FUNCTION_BLOCK FB_CartonCell EXTENDS SPT_BaseTypes.FB_PackML_BaseModule
VAR
    Line : FB_ContinuousLine;
    LineEvents : FB_LineEvents;
    Devices : FB_CellDevices;
    Stations : ARRAY[1..5] OF FB_StrokeStation;
    ActiveStation : DINT;
    Finished : BOOL;
    Cartons : DINT;
    AirFault : BOOL;
    LowStock : BOOL;
    PreviousState : Tc3_PackML_V2.E_PMLState;
    ActingScans : INT;
    RequestSample : DINT;
    Acknowledged : DINT;
    Accepted : BOOL;
    StatusBuffer : ARRAY[0..105] OF DINT;
END_VAR

METHOD PROTECTED Initialize : BOOL
// User mode 4 keeps Idle and Complete for one-station commissioning.
CustomModes(eMode := 4, sName := 'Manual stroke', bDisableHeld := TRUE,
    bDisableSuspended := TRUE, bEnableUnitModeChangeStopped := TRUE);
Initialize := SUPER^.Initialize();
END_METHOD

METHOD RunScan
IF _InitComplete THEN
    CyclicLogic();
ELSE
    _InitComplete := Initialize();
END_IF
END_METHOD

METHOD CyclicLogic
// SPT can call this hook while Initialize is still on the stack.
IF NOT _InitComplete THEN RETURN; END_IF

IF _CurrentState <> PreviousState THEN
    ActingScans := 0;
    PreviousState := _CurrentState;
ELSE
    ActingScans := MIN(45, ActingScans + 1);
END_IF

// Sample once so a concurrent ADS write belongs entirely to one scan.
RequestSample := GVL_HMI.Request;
IF RequestSample <> Acknowledged THEN
    Accepted := ApplyCommand(RequestSample MOD 256);
    Acknowledged := RequestSample;
END_IF

Line.Clock((_CurrentState = Tc3_PackML_V2.E_PMLState.ePMLState_Execute) AND Line.Enabled AND (_CurrentMode = E_PMLUnitMode.ePMLUnitMode_Production));
SUPER^.CyclicLogic();
LineEvents(Occurrence := Line.Occurrence, Alarm := Line.Alarm, Jammed := Line.Jammed,
    Idle := _CurrentState = Tc3_PackML_V2.E_PMLState.ePMLState_Idle);
PublishStatus();
END_METHOD

METHOD PROTECTED Execute
IF Line.Enabled AND (_CurrentMode = E_PMLUnitMode.ePMLUnitMode_Production) THEN
    IF Line.Alarm = 0 THEN Line.Step(Devices.MissingSeal); END_IF
    IF Line.Alarm <> 0 THEN ChangeState(Tc3_PackML_V2.E_PMLCommand.ePMLCommand_Abort); END_IF
    RETURN;
END_IF
IF (ActiveStation < 1) OR (ActiveStation > 5) THEN RETURN; END_IF
IF Finished THEN
    StateComplete();
    RETURN;
END_IF

Stations[ActiveStation].Step();
IF _CurrentMode = E_PMLUnitMode.ePMLUnitMode_Production THEN
    Devices.ProcessStation(ActiveStation, Stations[ActiveStation].Phase);
END_IF

IF Stations[ActiveStation].Done AND
   ((_CurrentMode = E_PMLUnitMode.ePMLUnitMode_UserMode1) OR Devices.ReadyToLeave(ActiveStation)) THEN
    IF (_CurrentMode = E_PMLUnitMode.ePMLUnitMode_UserMode1) OR (ActiveStation = 5) THEN
        Finished := TRUE;
        IF _CurrentMode = E_PMLUnitMode.ePMLUnitMode_Production THEN
            IF Devices.FinishCarton() THEN
                Cartons := Cartons + 1;
            END_IF
        END_IF
        StateComplete();
    ELSIF Devices.IndexToNext(ActiveStation) THEN
        ActiveStation := ActiveStation + 1;
    END_IF
END_IF
END_METHOD

METHOD PROTECTED Resetting
VAR
    StationIndex : INT;
END_VAR
FOR StationIndex := 1 TO 5 DO
    Stations[StationIndex].ResetStation();
END_FOR
Devices.ResetDevices();
Line.ResetLine();
ActiveStation := 0;
Finished := FALSE;
IF (_CurrentState = PreviousState) AND (ActingScans >= 45) THEN
    StateComplete();
END_IF
END_METHOD

METHOD PROTECTED Clearing
IF (_CurrentState = PreviousState) AND (ActingScans >= 45) THEN
    StateComplete();
END_IF
END_METHOD

METHOD PROTECTED Starting
IF (_CurrentState = PreviousState) AND (ActingScans >= 45) THEN
    StateComplete();
END_IF
END_METHOD

METHOD PROTECTED Stopping
IF (_CurrentState = PreviousState) AND (ActingScans >= 45) THEN
    StateComplete();
END_IF
END_METHOD

METHOD PROTECTED Aborting
IF (_CurrentState = PreviousState) AND (ActingScans >= 45) THEN
    StateComplete();
END_IF
END_METHOD

METHOD PROTECTED Holding
IF (_CurrentState = PreviousState) AND (ActingScans >= 45) THEN
    StateComplete();
END_IF
END_METHOD

METHOD PROTECTED Unholding
IF (_CurrentState = PreviousState) AND (ActingScans >= 45) THEN
    StateComplete();
END_IF
END_METHOD

METHOD PROTECTED Suspending
IF (_CurrentState = PreviousState) AND (ActingScans >= 45) THEN
    StateComplete();
END_IF
END_METHOD

METHOD PROTECTED Unsuspending
IF (_CurrentState = PreviousState) AND (ActingScans >= 45) THEN
    StateComplete();
END_IF
END_METHOD

METHOD PROTECTED Completing
IF (_CurrentState = PreviousState) AND (ActingScans >= 45) THEN
    StateComplete();
END_IF
END_METHOD

METHOD PRIVATE ApplyCommand : BOOL
VAR_INPUT
    Code : DINT;
END_VAR
VAR
    IsManual : BOOL;
END_VAR
IsManual := _CurrentMode = E_PMLUnitMode.ePMLUnitMode_UserMode1;
CASE Code OF
    E_ConsoleCommand.Reset:
        IF NOT AirFault AND ((_CurrentState = Tc3_PackML_V2.E_PMLState.ePMLState_Stopped) OR (_CurrentState = Tc3_PackML_V2.E_PMLState.ePMLState_Complete)) THEN
            ChangeState(Tc3_PackML_V2.E_PMLCommand.ePMLCommand_Reset);
            ApplyCommand := TRUE;
        END_IF
    E_ConsoleCommand.Start:
        IF NOT IsManual AND (_CurrentState = Tc3_PackML_V2.E_PMLState.ePMLState_Idle) THEN
            Line.Timing := Line.Enabled;
            ActiveStation := SEL(Line.Enabled, 1, 0);
            ChangeState(Tc3_PackML_V2.E_PMLCommand.ePMLCommand_Start);
            ApplyCommand := TRUE;
        END_IF
    E_ConsoleCommand.Hold:
        IF NOT IsManual AND (_CurrentState = Tc3_PackML_V2.E_PMLState.ePMLState_Execute) THEN
            ChangeState(Tc3_PackML_V2.E_PMLCommand.ePMLCommand_Hold);
            ApplyCommand := TRUE;
        END_IF
    E_ConsoleCommand.Unhold:
        IF _CurrentState = Tc3_PackML_V2.E_PMLState.ePMLState_Held THEN
            ChangeState(Tc3_PackML_V2.E_PMLCommand.ePMLCommand_Unhold);
            ApplyCommand := TRUE;
        END_IF
    E_ConsoleCommand.Suspend:
        IF NOT IsManual AND (_CurrentState = Tc3_PackML_V2.E_PMLState.ePMLState_Execute) THEN
            ChangeState(Tc3_PackML_V2.E_PMLCommand.ePMLCommand_Suspend);
            ApplyCommand := TRUE;
        END_IF
    E_ConsoleCommand.Unsuspend:
        IF _CurrentState = Tc3_PackML_V2.E_PMLState.ePMLState_Suspended THEN
            ChangeState(Tc3_PackML_V2.E_PMLCommand.ePMLCommand_Unsuspend);
            ApplyCommand := TRUE;
        END_IF
    E_ConsoleCommand.Stop:
        IF (_CurrentState <> Tc3_PackML_V2.E_PMLState.ePMLState_Undefined) AND
            (_CurrentState <> Tc3_PackML_V2.E_PMLState.ePMLState_Stopped) AND
            (_CurrentState <> Tc3_PackML_V2.E_PMLState.ePMLState_Stopping) AND
            (_CurrentState <> Tc3_PackML_V2.E_PMLState.ePMLState_Aborted) AND
            (_CurrentState <> Tc3_PackML_V2.E_PMLState.ePMLState_Aborting) AND
            (_CurrentState <> Tc3_PackML_V2.E_PMLState.ePMLState_Clearing) THEN
            Line.Timing := FALSE;
            ChangeState(Tc3_PackML_V2.E_PMLCommand.ePMLCommand_Stop);
            ApplyCommand := TRUE;
        END_IF
    E_ConsoleCommand.Abort:
        IF (_CurrentState <> Tc3_PackML_V2.E_PMLState.ePMLState_Aborted) AND
            (_CurrentState <> Tc3_PackML_V2.E_PMLState.ePMLState_Aborting) AND
            (_CurrentState <> Tc3_PackML_V2.E_PMLState.ePMLState_Undefined) THEN
            ChangeState(Tc3_PackML_V2.E_PMLCommand.ePMLCommand_Abort);
            ApplyCommand := TRUE;
        END_IF
    E_ConsoleCommand.Clear:
        IF NOT AirFault AND ((Line.Alarm = 0) OR ((Line.Alarm = 2) AND NOT Line.Jammed)) AND (_CurrentState = Tc3_PackML_V2.E_PMLState.ePMLState_Aborted) THEN
            Line.ClearAlarm();
            ChangeState(Tc3_PackML_V2.E_PMLCommand.ePMLCommand_Clear);
            ApplyCommand := TRUE;
        END_IF
    E_ConsoleCommand.Manual, E_ConsoleCommand.Automatic:
        IF _CurrentState = Tc3_PackML_V2.E_PMLState.ePMLState_Stopped THEN
            IF (Code = E_ConsoleCommand.Manual) AND NOT IsManual THEN
                Line.Timing := FALSE;
                ChangeMode(E_PMLUnitMode.ePMLUnitMode_UserMode1);
                ApplyCommand := TRUE;
            ELSIF (Code = E_ConsoleCommand.Automatic) AND IsManual THEN
                ChangeMode(E_PMLUnitMode.ePMLUnitMode_Production);
                ApplyCommand := TRUE;
            END_IF
        END_IF
    E_ConsoleCommand.Stroke1..E_ConsoleCommand.Stroke5:
        IF IsManual AND (_CurrentState = Tc3_PackML_V2.E_PMLState.ePMLState_Idle) THEN
            ActiveStation := Code - E_ConsoleCommand.Stroke1 + 1;
            ChangeState(Tc3_PackML_V2.E_PMLCommand.ePMLCommand_Start);
            ApplyCommand := TRUE;
        END_IF
    E_ConsoleCommand.DropAir:
        ApplyCommand := NOT AirFault;
        AirFault := TRUE;
        IF (_CurrentState <> Tc3_PackML_V2.E_PMLState.ePMLState_Aborted) AND (_CurrentState <> Tc3_PackML_V2.E_PMLState.ePMLState_Aborting) THEN
            ChangeState(Tc3_PackML_V2.E_PMLCommand.ePMLCommand_Abort);
        END_IF
    E_ConsoleCommand.RestoreAir:
        ApplyCommand := AirFault;
        AirFault := FALSE;
    E_ConsoleCommand.LowBlanks:
        ApplyCommand := NOT LowStock;
        LowStock := TRUE;
    E_ConsoleCommand.MissingSeal:
        ApplyCommand := NOT Devices.MissingSeal;
        Devices.MissingSeal := TRUE;
    E_ConsoleCommand.RestoreSeal:
        ApplyCommand := Devices.MissingSeal;
        Devices.MissingSeal := FALSE;
    E_ConsoleCommand.LoopLine, E_ConsoleCommand.Bench:
        IF NOT IsManual AND (_CurrentState = Tc3_PackML_V2.E_PMLState.ePMLState_Stopped) THEN
            ApplyCommand := Line.Enabled <> (Code = E_ConsoleCommand.LoopLine);
            Line.Timing := FALSE;
            Line.Enabled := Code = E_ConsoleCommand.LoopLine;
        END_IF
    E_ConsoleCommand.Standard, E_ConsoleCommand.Precision:
        IF Line.Enabled AND NOT IsManual AND (_CurrentState = Tc3_PackML_V2.E_PMLState.ePMLState_Stopped) THEN
            ApplyCommand := Line.Precision <> (Code = E_ConsoleCommand.Precision);
            Line.Precision := Code = E_ConsoleCommand.Precision;
        END_IF
    E_ConsoleCommand.JamClamp:
        IF Line.Enabled AND NOT IsManual AND NOT Line.Jammed AND (Line.Alarm = 0) THEN
            Line.Jammed := TRUE; ApplyCommand := TRUE;
        END_IF
    E_ConsoleCommand.ReleaseClamp:
        ApplyCommand := Line.Jammed; Line.Jammed := FALSE;
    E_ConsoleCommand.AckClamp:
        IF (_CurrentState = Tc3_PackML_V2.E_PMLState.ePMLState_Aborted) AND
            (Line.Alarm = 1) AND (RequestSample / 256 = Line.Occurrence) THEN
            Line.AcknowledgeAlarm(); ApplyCommand := TRUE;
        END_IF
    E_ConsoleCommand.Refill:
        ApplyCommand := LowStock;
        LowStock := FALSE;
END_CASE
END_METHOD

METHOD PRIVATE PublishStatus
StatusBuffer[0] := 51003;
StatusBuffer[1] := TO_DINT(_CurrentState);
StatusBuffer[2] := BOOL_TO_DINT(_CurrentMode = E_PMLUnitMode.ePMLUnitMode_UserMode1);
StatusBuffer[3] := ActiveStation;
StatusBuffer[4] := 0;
IF (ActiveStation >= 1) AND (ActiveStation <= 5) THEN
    StatusBuffer[4] := Stations[ActiveStation].Phase;
END_IF
StatusBuffer[5] := Cartons;
StatusBuffer[6] := BOOL_TO_DINT(AirFault);
StatusBuffer[7] := BOOL_TO_DINT(LowStock);
StatusBuffer[8] := Acknowledged;
StatusBuffer[9] := (StatusBuffer[9] MOD 2000000000) + 1;
StatusBuffer[10] := BOOL_TO_DINT(Accepted);
Devices.Publish(StatusBuffer);
Line.Publish(StatusBuffer);
GVL_HMI.Status := StatusBuffer;
END_METHOD

END_FUNCTION_BLOCK

(* stored: Version 1.1.0.1, ProductVersion 3.1.4024.53
   POU FB_CartonCell: Id {52592E20-A431-4FDA-93CC-000000000026}
   Method Initialize: Id {52592E20-A431-4FDA-93CC-000000000011}
   Method RunScan: Id {B9F992C3-0299-4AF4-A152-1426A98566B1}
   Method CyclicLogic: Id {52592E20-A431-4FDA-93CC-000000000012}
   Method Execute: Id {52592E20-A431-4FDA-93CC-000000000013}
   Method Resetting: Id {52592E20-A431-4FDA-93CC-000000000014}
   Method Clearing: Id {52592E20-A431-4FDA-93CC-000000000015}
   Method Starting: Id {52592E20-A431-4FDA-93CC-000000000016}
   Method Stopping: Id {52592E20-A431-4FDA-93CC-000000000017}
   Method Aborting: Id {52592E20-A431-4FDA-93CC-000000000018}
   Method Holding: Id {52592E20-A431-4FDA-93CC-000000000019}
   Method Unholding: Id {52592E20-A431-4FDA-93CC-000000000020}
   Method Suspending: Id {52592E20-A431-4FDA-93CC-000000000021}
   Method Unsuspending: Id {52592E20-A431-4FDA-93CC-000000000022}
   Method Completing: Id {52592E20-A431-4FDA-93CC-000000000023}
   Method ApplyCommand: Id {52592E20-A431-4FDA-93CC-000000000024}
   Method PublishStatus: Id {52592E20-A431-4FDA-93CC-000000000025} *)
